// TIA Portal project "PLC ile Tank Isıtıcı ve Mikser Otomasyonu" (V18)

(* hardware
DEVICE "S7-1200 station_1"  S7-1200 Station
   slot 0: "Rack_0"  S7-1200 Rack  Rack  V1.0
   slot 1: "PLC_1"  CPU 1214C DC/DC/Rly  6ES7 214-1HG40-0XB0  V4.6
*)

// ===== PLC "PLC_1"  CPU 1214C DC/DC/Rly =====

VAR_GLOBAL   // PLC tag table "Default tag table"
   "Start Butonu" AT %I0.0 : Bool;
   "Stop Butonu" AT %I0.1 : Bool;
   "Alt Seviye Sensörü" AT %I0.2 : Bool;
   "Üst Seviye Sensörü" AT %I0.3 : Bool;
   "PT100 Girişi" AT %IW96 : Int;
   "Isıtıcı" AT %Q0.0 : Bool;
   "Mikser" AT %Q0.1 : Bool;
   "Doldurma Valfi" AT %Q0.2 : Bool;
   "Boşaltma Valfi" AT %Q0.3 : Bool;
   "Sistem Genel Start" AT %M5.0 : Bool;
   "Tag_1" AT %MW20 : Int;
   "Tag_2" AT %MD22 : Real;
   "Sicaklik degeri" AT %MD26 : Real;
END_VAR

// folder: System blocks/Program resources

DATA_BLOCK "Timer-1"   // DB2
{ S7_Optimized_Access := 'TRUE' }
AUTHOR : Simatic
FAMILY : IEC
NAME : IEC_TMR
VERSION : 1.0
// stored: InstanceOfName IEC_TIMER
"IEC_TIMER"
BEGIN
END_DATA_BLOCK

// folder: (top level)

ORGANIZATION_BLOCK "Main"   // OB1, LAD, ProgramCycle
TITLE = "Main Program Sweep (Cycle)"
{ S7_Optimized_Access := 'TRUE' }
VERSION : 0.1
   VAR_INPUT
      Initial_Call : Bool;   // Initial call of this OB
      Remanence : Bool;   // =True, if remanent data are available
   END_VAR
BEGIN

REGION Network 1: SİSTEMİ BAŞLAT
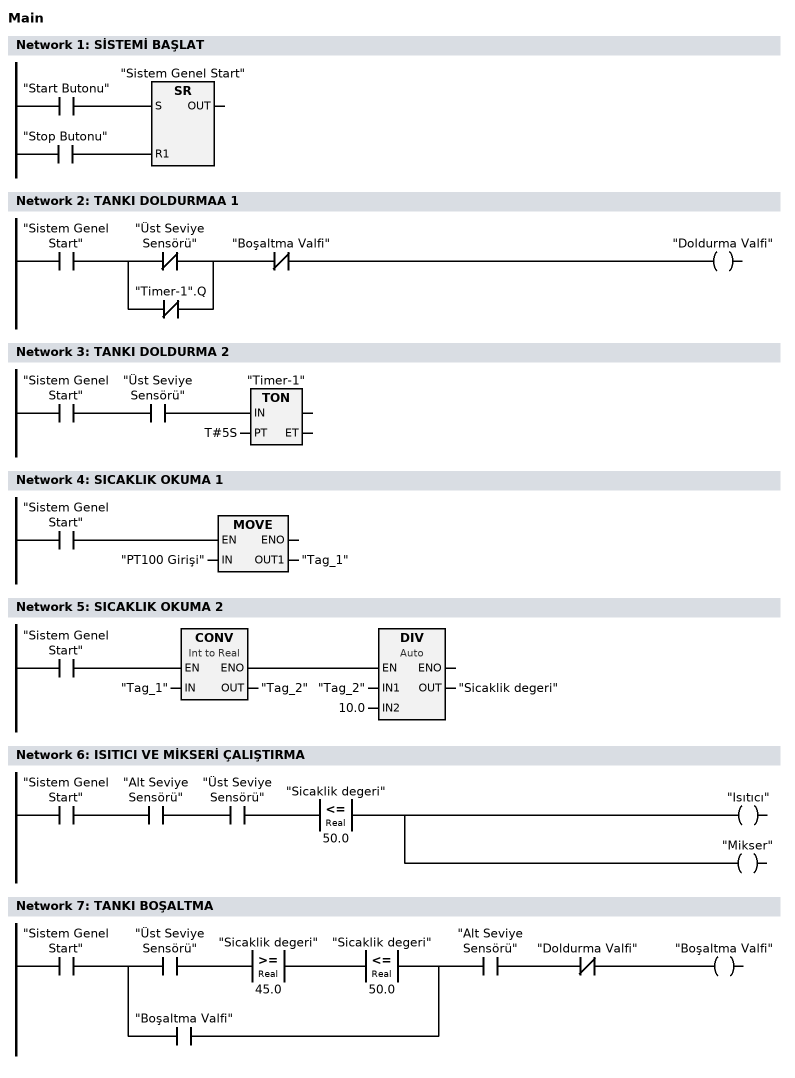
   RUNG wire#powerrail
      Contact( "Start Butonu" )
      S_SR(operand := "Sistem Genel Start", r1 := wire#w1)
   END_RUNG
   RUNG wire#powerrail
      Contact( "Stop Butonu" )
   END_RUNG wire#w1
   // the same network as SCL:
   IF "Start Butonu" THEN
       "Sistem Genel Start" := TRUE;   // SR flip-flop
   END_IF;
   IF "Stop Butonu" THEN "Sistem Genel Start" := FALSE; END_IF;
END_REGION

REGION Network 2: TANKI DOLDURMAA 1
   RUNG wire#powerrail
      Contact( "Sistem Genel Start" )
      wire#w1
      I_Contact( "Üst Seviye Sensörü" )
      wire#w2
      I_Contact( "Boşaltma Valfi" )
      Coil( "Doldurma Valfi" )
   END_RUNG
   RUNG wire#w1
      I_Contact( "Timer-1".Q )
   END_RUNG wire#w2
   // the same network as SCL:
   "Doldurma Valfi" := "Sistem Genel Start" AND (NOT "Üst Seviye Sensörü" OR NOT "Timer-1".Q) AND NOT "Boşaltma Valfi";
END_REGION

REGION Network 3: TANKI DOLDURMA 2
   "Timer-1".TON(IN := "Sistem Genel Start" AND "Üst Seviye Sensörü", PT := T#5S);
END_REGION

REGION Network 4: SICAKLIK OKUMA 1
   RUNG wire#powerrail
      Contact( "Sistem Genel Start" )
      Move(in := "PT100 Girişi", out1 => "Tag_1")
   END_RUNG
   // the same network as SCL:
   IF "Sistem Genel Start" THEN "Tag_1" := "PT100 Girişi"; END_IF;
END_REGION

REGION Network 5: SICAKLIK OKUMA 2
   RUNG wire#powerrail
      Contact( "Sistem Genel Start" )
      { S7_Templates := "[SrcType := Int, DestType := Real]" } Convert(in := "Tag_1", out => "Tag_2")
      Div(in1 := "Tag_2", in2 := 10.0, out => "Sicaklik degeri")
   END_RUNG
   // the same network as SCL:
   IF "Sistem Genel Start" THEN
       "Tag_2" := INT_TO_REAL("Tag_1");
       "Sicaklik degeri" := "Tag_2" / 10.0;
   END_IF;
END_REGION

REGION Network 6: ISITICI VE MİKSERİ ÇALIŞTIRMA
   RUNG wire#powerrail
      Contact( "Sistem Genel Start" )
      Contact( "Alt Seviye Sensörü" )
      Contact( "Üst Seviye Sensörü" )
      { S7_Templates := "SrcType := Real" } LE_Contact(in1 := "Sicaklik degeri", in2 := 50.0)
      wire#w1
      Coil( "Isıtıcı" )
   END_RUNG
   RUNG wire#w1
      Coil( "Mikser" )
   END_RUNG
   // the same network as SCL:
   "Isıtıcı" := "Sistem Genel Start" AND "Alt Seviye Sensörü" AND "Üst Seviye Sensörü" AND ("Sicaklik degeri" <= 50.0);
   "Mikser" := "Isıtıcı";
END_REGION

REGION Network 7: TANKI BOŞALTMA
   RUNG wire#powerrail
      Contact( "Sistem Genel Start" )
      wire#w1
      Contact( "Üst Seviye Sensörü" )
      { S7_Templates := "SrcType := Real" } GE_Contact(in1 := "Sicaklik degeri", in2 := 45.0)
      { S7_Templates := "SrcType := Real" } LE_Contact(in1 := "Sicaklik degeri", in2 := 50.0)
      wire#w2
      Contact( "Alt Seviye Sensörü" )
      I_Contact( "Doldurma Valfi" )
      Coil( "Boşaltma Valfi" )
   END_RUNG
   RUNG wire#w1
      Contact( "Boşaltma Valfi" )
   END_RUNG wire#w2
   // the same network as SCL:
   "Boşaltma Valfi" := "Sistem Genel Start" AND (("Üst Seviye Sensörü" AND ("Sicaklik degeri" >= 45.0) AND ("Sicaklik degeri" <= 50.0)) OR "Boşaltma Valfi") AND "Alt Seviye Sensörü" AND NOT "Doldurma Valfi";
END_REGION
END_ORGANIZATION_BLOCK